// TIA Portal V21 export
// export: Created 2026-11-21T13:24:05.0270368Z, ExportSetting WithDefaults, DisplayName Totally Integrated Automation Portal, DisplayVersion V21, DisplayName STEP 7 Professional, DisplayVersion V21, DisplayName STEP 7 Safety, DisplayVersion V21, DisplayName Tech WebApplication, DisplayVersion V21, DisplayName WinCC Basic/Comfort/Advanced, DisplayVersion V21, DisplayName WinCC Unified, DisplayVersion V21
FUNCTION_BLOCK "LockedSafety"   // FB1, F_FBD
{ S7_Optimized_Access := 'TRUE' }
VERSION : 0.1
// Main safety block of a safety program with a password.
// stored: AutoNumber true, IsIECCheckEnabled false, UDAEnableTagReadback false
   VAR
      source : Bool;
      target : Bool;
   END_VAR
BEGIN

REGION Network 1: Copy
   // Copies one bit to another.
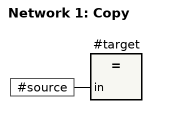
   #target := #source;
END_REGION
END_FUNCTION_BLOCK
